PROGRAM prg_InterCon_Usage
VAR
END_VAR

// TriBlender  

IF fbElement[E_Element_List.eTank_1].eState_Short=E_Element_State_Short.eClean 
AND fbElement[E_Element_List.eTriBlender_Marinada].eState_Short=E_Element_State_Short.eClean
THEN;
	//eIntCon_TriB_T1_Marin:=E_InterConnection.Avalable;
END_IF

act_Call_InterConnection();

CASE eTriBlenderUsage OF
	E_TriBlenderUsage.eMarinada_T1,E_TriBlenderUsage.eMarinada_T2:;
		fbElement[E_Element_List.eTriBlender_Marinada].m_StateUpdate_Limit(value:=TRUE);		
		fbElement[E_Element_List.eTriBlender_Color].m_StateUpdate_Limit(value:=TRUE);
	
	E_TriBlenderUsage.eMarinada_Standby:;
		fbElement[E_Element_List.eTriBlender_Marinada].m_StateUpdate_Limit(value:=FALSE);
		fbElement[E_Element_List.eTriBlender_Color].m_StateUpdate_Limit(value:=TRUE);
		
	E_TriBlenderUsage.eColor_T3,E_TriBlenderUsage.eColor_T4:;	
		fbElement[E_Element_List.eTriBlender_Marinada].m_StateUpdate_Limit(value:=TRUE);		
		fbElement[E_Element_List.eTriBlender_Color].m_StateUpdate_Limit(value:=TRUE);
	
	E_TriBlenderUsage.eColor_Standby:;	
		fbElement[E_Element_List.eTriBlender_Marinada].m_StateUpdate_Limit(value:=TRUE);
		fbElement[E_Element_List.eTriBlender_Color].m_StateUpdate_Limit(value:=FALSE);
ELSE;
		fbElement[E_Element_List.eTriBlender_Marinada].m_StateUpdate_Limit(value:=FALSE);
		fbElement[E_Element_List.eTriBlender_Color].m_StateUpdate_Limit(value:=FALSE);	
END_CASE

CASE ePrL_M_Usage OF
	E_PrLine_M_LineUsage.eMarinada_T1,
	E_PrLine_M_LineUsage.eMarinada_T2:;
		fbElement[E_Element_List.eLine_Marinada].m_StateUpdate_Limit(value:=TRUE);
	E_PrLine_M_LineUsage.eNotInUse:;
		fbElement[E_Element_List.eLine_Marinada].m_StateUpdate_Limit(value:=FALSE);
END_CASE

CASE ePrL_C_Usage OF
	E_PrLine_C_Usage.eColor_T3,
	E_PrLine_C_Usage.eColor_T4:;
		fbElement[E_Element_List.eLine_Color].m_StateUpdate_Limit(value:=TRUE);
	E_PrLine_C_Usage.eNotInUse:;
		fbElement[E_Element_List.eLine_Color].m_StateUpdate_Limit(value:=FALSE);
END_CASE
(*
IF eTriBlenderPipe_In=eTriBlenderPipe_Out THEN;
	eTriBlenderPipe:=eTriBlenderPipe_In;
ELSE;
	eTriBlenderPipe:=E_TriBlenderPipe.eNone;
END_IF
*)
(*
CASE fbTriBlender_Select.eStatus OF
	E_TriBlenderSelect.eMarinade:;
		eTriBlenderPipe:=E_TriBlenderPipe.eMarinada;	
	E_TriBlenderSelect.eColor:;
		eTriBlenderPipe:=E_TriBlenderPipe.eColor;
	E_TriBlenderSelect.eDrain:;
		eTriBlenderPipe:=E_TriBlenderPipe.eNone;
ELSE;
	eTriBlenderPipe:=E_TriBlenderPipe.eNone;	
END_CASE
*)

ACTION act_Call_InterConnection:
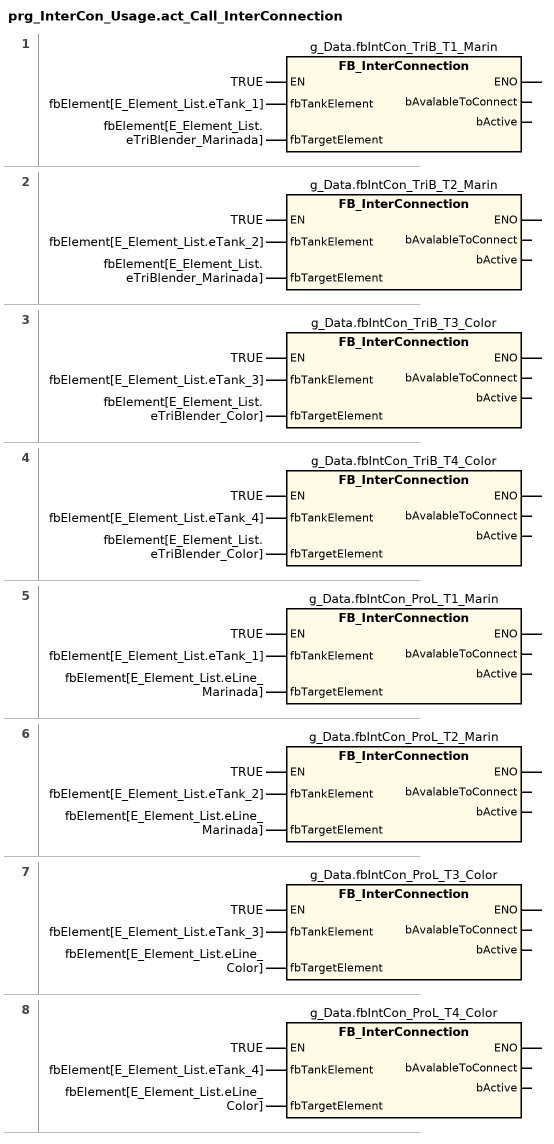
// NETWORK 1
g_Data.fbIntCon_TriB_T1_Marin(fbTankElement := fbElement[E_Element_List.eTank_1], fbTargetElement := fbElement[E_Element_List.eTriBlender_Marinada]); // FB_InterConnection

// NETWORK 2
g_Data.fbIntCon_TriB_T2_Marin(fbTankElement := fbElement[E_Element_List.eTank_2], fbTargetElement := fbElement[E_Element_List.eTriBlender_Marinada]); // FB_InterConnection

// NETWORK 3
g_Data.fbIntCon_TriB_T3_Color(fbTankElement := fbElement[E_Element_List.eTank_3], fbTargetElement := fbElement[E_Element_List.eTriBlender_Color]); // FB_InterConnection

// NETWORK 4
g_Data.fbIntCon_TriB_T4_Color(fbTankElement := fbElement[E_Element_List.eTank_4], fbTargetElement := fbElement[E_Element_List.eTriBlender_Color]); // FB_InterConnection

// NETWORK 5
g_Data.fbIntCon_ProL_T1_Marin(fbTankElement := fbElement[E_Element_List.eTank_1], fbTargetElement := fbElement[E_Element_List.eLine_Marinada]); // FB_InterConnection

// NETWORK 6
g_Data.fbIntCon_ProL_T2_Marin(fbTankElement := fbElement[E_Element_List.eTank_2], fbTargetElement := fbElement[E_Element_List.eLine_Marinada]); // FB_InterConnection

// NETWORK 7
g_Data.fbIntCon_ProL_T3_Color(fbTankElement := fbElement[E_Element_List.eTank_3], fbTargetElement := fbElement[E_Element_List.eLine_Color]); // FB_InterConnection

// NETWORK 8
g_Data.fbIntCon_ProL_T4_Color(fbTankElement := fbElement[E_Element_List.eTank_4], fbTargetElement := fbElement[E_Element_List.eLine_Color]); // FB_InterConnection
END_ACTION

END_PROGRAM

(* stored: Version 1.1.0.1, ProductVersion 3.1.4024.13
   POU prg_InterCon_Usage: Id {24fec81d-d792-4666-bec4-7cc918d6b551}, SpecialFunc None
   Action act_Call_InterConnection: Id {f183bb8e-cf96-4bd4-ba1b-976dcd989a9c} *)
